TYPE T_SetConfigParamList : ARRAY[1..Param_Config.MaxConfigParamPerModule] OF ST_SetConfigParamParam;
END_TYPE

(* stored: Version 1.1.0.1, ProductVersion 3.1.4026.18
   DUT T_SetConfigParamList: Id {ee14efc3-2972-48df-98dd-a170adca18c3} *)
